// TIA Portal V19 export
TYPE "ST_Reset"
   STRUCT
      Execute : Bool;
      Busy : Bool;
      Done : Bool;
      Error : Bool;
      ErrorID : Word;
   END_STRUCT;
END_TYPE
